(* IEC 61131-3 sources: avi-aoi-management/scripts/ai-eval/ngau-nhien/kho/st-tv2-dem-san-pham/khung/src, 1 file *)

(* ---- DemSanPham.st ---- *)
FUNCTION_BLOCK DemSanPham
VAR_INPUT
    CAM_BIEN : BOOL;
    KICH_THUOC_LO : INT;
    RESET : BOOL;
END_VAR
VAR_OUTPUT
    DEM : INT;
    XONG_LO : BOOL;
    SO_LO : INT;
END_VAR
    (* TODO: cài đặt theo đề bài, dùng R_TRIG + CTU *)
    DEM := 0;
END_FUNCTION_BLOCK
